Fanuc KAREL source: KT00679.KL

PROGRAM KT00679
%NOLOCKGROUP
VAR
  P1: JOINTPOS
  P2: JOINTPOS
  OUT: INTEGER
BEGIN
  OUT = NOT P1
END KT00679
